TYPE ST_AlarmIn :
STRUCT
	arbFatalError			:ARRAY[0..nALARM_MAX_NO] OF ST_AlarmProperties;
	arbError				:ARRAY[0..nALARM_MAX_NO] OF ST_AlarmProperties;
	arbWarning			:ARRAY[0..nALARM_MAX_NO] OF ST_AlarmProperties;
	arbMessage			:ARRAY[0..nALARM_MAX_NO] OF ST_AlarmProperties;
	arbHint				:ARRAY[0..nALARM_MAX_NO] OF ST_AlarmProperties;
END_STRUCT
END_TYPE

(* stored: Version 1.1.0.1, ProductVersion 3.1.4024.15
   DUT ST_AlarmIn: Id {5fd51be2-c57e-46e8-a43c-bebda06f1c70} *)
